FUNCTION F_ConvArrBitsToWord : WORD
VAR_INPUT
	arrBits: ARRAY [0..15] OF BOOL;
END_VAR
VAR
END_VAR

F_ConvArrBitsToWord := 0;

END_FUNCTION

(* stored: Version 1.1.0.1, ProductVersion 3.1.4024.15
   POU F_ConvArrBitsToWord: Id {70052612-e166-4544-872b-d6a6e3a99fa1}, SpecialFunc None *)
